TYPE "G003_type"
TITLE = %version: 5.09 % %Commit:  c3808b61 % CN: 10
VERSION : 0.1
//
//SOURCE
//%Project:      allcttt %
//%Repo:         a_ttt %
//%Commit:       c3808b61 %
//%DateTimeUTC:  2023-12-11T14:59:55 %
//
//%HISTORY%
//Issue:        Commit:  Date:      Version: Author:              Description:
//------------- -------- ---------- -------- -------------------- ------------------------------------------------------------------------------
//ALLCTTT-4059  c3808b61 2023-12-11 5.09     Pascal van Kempen    Added history table
//ALLCTTT-4042  55fd833f 2023-12-05 5.08     Henri de Leijer      First step to remove the library files
//ALLCTTT-1873  b29a070d 2022-03-17 5.07     Henri de Leijer      ALLCTTT-1873 TB08 of HSZ51 report PEC blockage error
//ALLCTTT-272   544e4e84 2020-12-10 5.06     Pascal van Kempen    removed keywords
//ALLCTTT-272   9d531fbf 2020-12-10 5.05     Pascal van Kempen    Revert corrected checkin sequence for determining version information properly
//ALLCTTT-272   ae3fa862 2020-12-10 5.04     Pascal van Kempen    corrected checkin sequence for determining version information properly
//ALLCTTT-272   5a1edb78 2020-12-10 5.03     Pascal van Kempen    Revert keywords updates
//ALLCTTT-272   8d62c219 2020-12-10 5.02     Pascal van Kempen    keywords updates
//ALLCTTT-272   31a64871 2020-12-10 5.01     Pascal van Kempen    initial import
//
//Modification History:                                 By:      Date:     Rev:
//----------------------------------------------------  -------  --------  -----
//Initial version                                       nlHdL    07-01-20   2.01
   STRUCT
      OBT_onto_HSZ : Bool;   //Command signal from ACZ to HSZ and DCZ that OBT is entering High Speed
      HSZ_Stop_Req : Bool;   //Request signal from HSZ to DCZ that section has stop request
      DCZ_Halt_Die_Back : Bool;   //Command signal from DCZ to halt section in Die-Back
      Spare_0_3 : Bool;   //Spare_0_3
      Spare_0_4 : Bool;   //Spare_0_4
      Spare_0_5 : Bool;   //Spare_0_5
      Spare_0_6 : Bool;   //Spare_0_6
      Spare_0_7 : Bool;   //Spare_0_7
      Spare_1_0 : Bool;   //Spare_1_0
      Spare_1_1 : Bool;   //Spare_1_1
      Spare_1_2 : Bool;   //Spare_1_2
      Spare_1_3 : Bool;   //Spare_1_3
      Spare_1_4 : Bool;   //Spare_1_4
      Spare_1_5 : Bool;   //Spare_1_5
      Spare_1_6 : Bool;   //Spare_1_6
      Spare_1_7 : Bool;   //Spare_1_7
      Cascade_Delay_Time : Int;   //  [ms] Cascade delay time
   END_STRUCT;

END_TYPE
